(* IEC 61131-3 sources: PLC-Static-Analysis/modules/plc-rules/src/test/resources/PLCA-Q014/allowed, 1 file *)

(* ---- a.st ---- *)
FUNCTION F_Scale : REAL
VAR_INPUT
    r : REAL;
END_VAR
F_Scale := r * 3.6 + 273.15; // PLCA-Q014
END_FUNCTION
